Staubli VAL3: saveTRAJ.dtx

public trajItem tTrajItem{}
  [Key1]
    pointItem pPointItem
      [0]
        paraItem pParaItem
          [0]
            mdesc mMdesc
            num nMoveType
            num nActionIndex[2]
            num nPercentage[2]
        pointRx pPointRx
        jointRx jJointRx
    num nFrameIndex
    num nToolIndex
    string sID
    num nMoveID
